{attribute 'qualified_only'}
{attribute 'strict'}
TYPE E_CheckMagazines_New :
(
	eIdle	:= 0,
	eStartNewNCI	:= 1,
	eDebug := 2,
	eWaitForPortal := 3
);
END_TYPE

(* stored: Version 1.1.0.1, ProductVersion 3.1.4024.12
   DUT E_CheckMagazines_New: Id {6fb68d0d-96e3-4d3b-8bbf-a2242f2f2e7c} *)
